Fanuc KAREL source: KC00064.KL

PROGRAM KC00064
%NOLOCKGROUP
%ENVIRONMENT CVIS
VAR
  I: INTEGER
  J: INTEGER
  K: INTEGER
  R: REAL
  B: BOOLEAN
  S: STRING[80]
  T: STRING[80]
  P: PATH
  Q: PATH
  AI: ARRAY[8] OF INTEGER
  AB: ARRAY[244] OF BYTE
BEGIN
  V_INIT_QUEUE(I,J)
END KC00064
